Fanuc KAREL source: KT00762.KL

PROGRAM KT00762
%NOLOCKGROUP
VAR
  R1: REAL
  R2: REAL
  OUT: INTEGER
BEGIN
  R1 = 2.0
  R2 = 3.0
  R1 = 2.0
  R2 = 3.0
  OUT = ACOS(R1)
END KT00762
